(* CODESYS project xy_plotter.export

Project tree, tasks and I/O mapping:
  Device : CODESYS Control for Raspberry Pi 64 SL, CODESYS, order no. 2302000009, version 4.21.0.0
    application Application
      libraries: Standard, 3.5.22.0 (System); Net Base Services, * (CODESYS)
      task Main_OB1 (cyclic, interval t#4ms, priority 1) calls FB100_Logic_Call
      Drawing/
        global variables Drawing
      ESP Data/
        global variables RCV_ESP_Buffer
        global variables SND_ESP_Buffer
      HMI Data/
        global variables DB
      PLC data types/
        data type ESP_Cmd
        data type ESP_Coord
        data type ESP_Resp
        data type ESP_Zsw
        data type PLC_Contour
        data type PLC_Point
        data type TMR
        TCP/
          data type TCP_Con
          data type TCP_ESP_RCV
          data type TCP_ESP_SND
          data type TCP_Rcv
          data type TCP_Snd
      program FB100_Logic_Call [ST]
      function block FB200_TCP_ESP [ST]
      function block FB300_ESP_Cmd [ST]: AssignBit
      Symbols
    SoftMotion General Axis Pool
    GPIOs_A_B : GPIOs A/B, CODESYS, version 4.21.0.0
        unmapped channels: digital inputs (GPIO0..GPIO31), digital outputs (GPIO0..GPIO31)
    Onewire
    Camera device
      <Empty>
    SPI
    I²C
*)

// Device/Application/PLC data types/ESP_Cmd
TYPE ESP_Cmd :
	
STRUCT
    Stw         : UINT := 0;   // ESP32 control word
    PointFlags  : UINT := 0;   // Point command flags
    ContourNum  : UINT := 0;   // Contour number
    PointNum    : UINT := 0;   // Point number
    Speed       : UINT := 0;   // Movement speed
    Coord_X     : UINT := 0;   // Target X coordinate
    Coord_Y     : UINT := 0;   // Target Y coordinate
	
	ManMoveSpeed		: UINT := 0;	// Manual movement speed	
	
	TargetX         	: UINT := 0;   // Target X coordinate
	TargetY         	: UINT := 0;   // Target Y coordinate
	TargetMoveSpeed 	: UINT := 0;   // Target movement speed
		
END_STRUCT

END_TYPE

// Device/Application/PLC data types/ESP_Coord
TYPE ESP_Coord :
	
STRUCT
    X : REAL := 0.0;
    Y : REAL := 0.0;
END_STRUCT

END_TYPE

// Device/Application/PLC data types/ESP_Resp
TYPE ESP_Resp :

STRUCT
    ZSW_Byte1     : BYTE := 16#00;      // Status byte 1
    ZSW_Byte2     : BYTE := 16#00;      // Status byte 2
    NumExpected   : UINT := 0;          // Next expected point number
    LastContRcv   : UINT := 0;          // Last contour received
    LastContDone  : UINT := 0;          // Last contour completed
    CurrPoint     : UINT := 0;          // Current point number
    Coord_X       : UINT := 0;          // Current X coordinate
    Coord_Y       : UINT := 0;          // Current Y coordinate
    PointsInBuffer: UINT := 0;          // Number of points currently stored
    ErrorCode     : UINT := 0;          // ESP32 error code
	DrawingState  : USINT := 0;	    	// Running - 1, aborted - 2, finished - 3
END_STRUCT

END_TYPE

// Device/Application/PLC data types/ESP_Zsw
TYPE ESP_Zsw :
	
STRUCT
    RdyForRcvNewPnt 	: BOOL := FALSE;
    RdyForEn        	: BOOL := FALSE;
    Enabled         	: BOOL := FALSE;
    Off1            	: BOOL := FALSE;
    Off2            	: BOOL := FALSE;
    PenDn           	: BOOL := FALSE;
    RdyStartNewDrw  	: BOOL := FALSE;
    RdyContPrevDrw  	: BOOL := FALSE;
    DrwProccAct     	: BOOL := FALSE;
    SnsrHomeX       	: BOOL := FALSE;
    SnsrHomeY       	: BOOL := FALSE;
    SnsrLimitX      	: BOOL := FALSE;
    SnsrLimitY      	: BOOL := FALSE;
    MovingAuto      	: BOOL := FALSE;
    MovingHome      	: BOOL := FALSE;
    MovingManual    	: BOOL := FALSE;
END_STRUCT

END_TYPE

// Device/Application/PLC data types/PLC_Contour
TYPE PLC_Contour :

STRUCT
    RcvdByEsp    : BOOL := FALSE;   // Contour received by ESP32
    Done         : BOOL := FALSE;   // Contour drawing completed
    StartIndex   : UINT := 0;       // Start index of contour in point buffer
    PointCount   : UINT := 0;       // Number of points in contour
    CurrentPoint : UINT := 0;       // Current point number
END_STRUCT

END_TYPE

// Device/Application/PLC data types/PLC_Point
TYPE PLC_Point :
	
STRUCT
    CmdType : UINT := 0;     // Point command type
    Speed   : UINT := 0;     // Movement speed
    Coord_X : UINT := 0;     // Target X coordinate
    Coord_Y : UINT := 0;     // Target Y coordinate
END_STRUCT

END_TYPE

// Device/Application/PLC data types/TMR
TYPE TMR :

STRUCT
	IN : BOOL := FALSE;      // Timer enable input
    PT : TIME := T#0MS;      // Preset time
    Q  : BOOL := FALSE;      // Timer output
END_STRUCT

END_TYPE

// Device/Application/PLC data types/TCP/TCP_Con
TYPE TCP_Con :

STRUCT
    Req    		: BOOL;
    Done   		: BOOL;
    Busy   		: BOOL;
    Error  		: BOOL;
	ErrorID		: NBS.ERROR;
    Active		: BOOL;
	ConnBusy    : BOOL;
	ConnError   : BOOL;
	ConnErrorID : NBS.ERROR;
	Connected   : BOOL;
END_STRUCT

END_TYPE

// Device/Application/PLC data types/TCP/TCP_ESP_RCV
TYPE TCP_ESP_RCV :
	
STRUCT
	ResponseZswByte1       : BYTE;         		// ESP32 status word
	ResponseZswByte2       : BYTE;         		// ESP32 status word
    ResponseNumExpected    : UINT := 0;    		// Next expected point number
    ResponseLastContRcv    : UINT := 0;    		// Last contour received
    ResponseLastContDone   : UINT := 0;    		// Last contour completed
    ResponseCurrPoint      : UINT := 0;    		// Current point number
    ResponseCoord_X        : UINT := 0;   		// Current X coordinate
    ResponseCoord_Y        : UINT := 0;    		// Current Y coordinate
    ResponsePointsInBuffer : UINT := 0;    		// Number of points currently stored in buffer
    ResponseErrorCode      : UINT := 0;    		// ESP32 error code
	ResponseDrawingState   : USINT := 0;	    // Running - 1, aborted - 2, finished - 3
END_STRUCT

END_TYPE

// Device/Application/PLC data types/TCP/TCP_ESP_SND
TYPE TCP_ESP_SND :
	
STRUCT
	CommandStw        : UINT := 0;   			// ESP32 control word
    CommandPointFlags : UINT := 0;   			// Point command flags
    CommandContourNum : UINT := 0;   			// Contour number
    CommandPointNum   : UINT := 0;   			// Point number
    CommandSpeed      : UINT := 0;   			// Movement speed
    CommandCoord_X    : UINT := 0;   			// Target X coordinate
    CommandCoord_Y    : UINT := 0;   			// Target Y coordinate
	CommandManMoveSpeed		: UINT := 0;		// Manual movement speed	
	CommandTargetX         	: UINT := 0;   		// Target X coordinate
	CommandTargetY         	: UINT := 0;   		// Target Y coordinate
	CommandTargetMoveSpeed 	: UINT := 0;   		// Target movement speed
END_STRUCT

END_TYPE

// Device/Application/PLC data types/TCP/TCP_Rcv
TYPE TCP_Rcv :

STRUCT
    Req    		: BOOL;
	Ndr    		: BOOL;
    Done   		: BOOL;
    Busy   		: BOOL;
    Error  		: BOOL;
	ErrorID		: NBS.ERROR;
    Status		: WORD;
	Len			: UDINT;
END_STRUCT

END_TYPE

// Device/Application/PLC data types/TCP/TCP_Snd
TYPE TCP_Snd :

STRUCT
    Req    		: BOOL;
    Done   		: BOOL;
    Busy   		: BOOL;
    Error  		: BOOL;
	ErrorID		: NBS.ERROR;
    Status		: WORD;
	Len			: UDINT;
END_STRUCT

END_TYPE

// Device/Application/Drawing/Drawing
{attribute 'qualified_only'}
VAR_GLOBAL
	
	TotalNumbContours 	: UINT := 0;                    	// Total number of contours
    TotalNumbPoints   	: UINT := 0;                    	// Total number of points

    Contour 			: ARRAY[0..700] OF PLC_Contour;     // Contour data array
    Points  			: ARRAY[0..7000] OF PLC_Point;      // Point data array

END_VAR

// Device/Application/ESP Data/RCV_ESP_Buffer
{attribute 'qualified_only'}
VAR_GLOBAL
	
    TCP_ESP_RCV	: TCP_ESP_RCV;         		

END_VAR

// Device/Application/ESP Data/SND_ESP_Buffer
{attribute 'qualified_only'}
VAR_GLOBAL
	TCP_ESP_SND : TCP_ESP_SND;
	Default : TCP_ESP_SND;
END_VAR

// Device/Application/HMI Data/DB
{attribute 'qualified_only'}
VAR_GLOBAL
	
    RcvDataFromPC : BOOL := FALSE; 					// Receive new data from PC												
    AutoCmd : BOOL := FALSE;						// Start automatic operation
    MoveCmd : BOOL := TRUE;							// Enable move
    HomeCmd : BOOL := FALSE;						// Start homing sequence
	MoveToTargetCmd : BOOL := FALSE;				// Start moving to target (during manual mode)
    StopCmd : BOOL := TRUE;							// Stop current operation
    EstopCmd : BOOL := FALSE;						// Emergency stop command
    CleanCmd : BOOL := FALSE;						// Clear ESP32 point buffer
    
	ManualPenDn : BOOL := FALSE;					// Move pen to down position manually
    ManMoveNorth : BOOL := FALSE;					// Manual movement commands
    ManMoveNEast : BOOL := FALSE;
    ManMoveEast  : BOOL := FALSE;
    ManMoveSEast : BOOL := FALSE;
    ManMoveSouth : BOOL := FALSE;
    ManMoveSWest : BOOL := FALSE;
    ManMoveWest  : BOOL := FALSE;
    ManMoveNWest : BOOL := FALSE;
	ManMoveSpeed : INT := 1000;
	
	TargetX : INT := 0;								 // Move to point (during manual mode)
	TargetY : INT := 0;
	TargetMoveSpeed : INT := 1000;
	TargetPenDn : BOOL := FALSE;
	
END_VAR

// Device/Application/FB100_Logic_Call
PROGRAM FB100_Logic_Call

VAR
	TcpPcDone      : BOOL := FALSE;
    TcpPcDataSaved : BOOL := FALSE;	

    xDeleteDrwReq  : BOOL := FALSE;
    xDeleteDrwDone : BOOL := FALSE;
    xAckReq        : BOOL := FALSE;
    xAckReset      : BOOL := FALSE;

    xEspConnected  : BOOL := FALSE;
    xEspSendDone   : BOOL := FALSE;
    xEspReceiveNdr : BOOL := FALSE;
    xEspSendReq    : BOOL := FALSE;
    xEspReceiveReq : BOOL := FALSE;

    xEspHomeX      : BOOL := FALSE;
    xEspHomeY      : BOOL := FALSE;
	
	PlcHeartbeat   : UDINT := 0;
	
	TargetReached  : BOOL := FALSE;
	
	EspCommLostTimer 	: TON;
	EspCommLost 		: BOOL := FALSE;
	
	FB300_ESP_Cmd : FB300_ESP_Cmd;
	FB200_TCP_ESP : FB200_TCP_ESP;
END_VAR

VAR CONSTANT
    RcvPcBufferSize : INT := 500;
    DrwContourSize  : INT := 500;
    DrwPointSize    : INT := 7000;
END_VAR


// pc: 192.168.0.100
// plc: 192.168.0.254
// esp: 192.168.0.154

// Plc Heartbit for Ignition
PlcHeartbeat := PlcHeartbeat + 2;

// Reset the homing command when automatic mode is active or both axes have reached their home positions
IF DB.AutoCmd OR (xEspHomeX AND xEspHomeY) THEN
	DB.HomeCmd := FALSE;
END_IF;

IF RCV_ESP_Buffer.TCP_ESP_RCV.ResponseLastContDone >= Drawing.TotalNumbContours THEN
	DB.AutoCmd := FALSE;
END_IF

// Reset the target moving command when both axes have reached their positions
TargetReached := ABS(UINT_TO_INT(RCV_ESP_Buffer.TCP_ESP_RCV.ResponseCoord_X) - DB.TargetX * 100) <= 1 AND ABS(UINT_TO_INT(RCV_ESP_Buffer.TCP_ESP_RCV.ResponseCoord_Y) - DB.TargetY * 100) <= 1;

IF DB.MoveToTargetCmd AND TargetReached THEN
    DB.MoveToTargetCmd := FALSE;
END_IF;

// Cancel automatic movement and homing when a stop command is active
IF DB.StopCmd THEN
	DB.AutoCmd := FALSE;
	DB.HomeCmd := FALSE;
	DB.MoveToTargetCmd := FALSE;
END_IF;

// Prepare commands and exchange drawing data with the ESP
FB300_ESP_Cmd(Enable := NOT DB.RcvDataFromPC,
              ContourTotalNum := Drawing.TotalNumbContours,
              PointsTotalNum := Drawing.TotalNumbPoints,
              TCP_Conn_Estab := xEspConnected,
              TCP_Snd_Done := xEspSendDone,
              TCP_Rcv_Ndr := xEspReceiveNdr,
			  ConnLost := EspCommLost,
              TCP_Snd_Req => xEspSendReq,
              TCP_Rcv_Req => xEspReceiveReq,
			  SnsrHomeX => xEspHomeX,
              SnsrHomeY => xEspHomeY);
			  
// Manage the TCP connection and data exchange between the PLC and ESP
FB200_TCP_ESP(Enable := NOT DB.RcvDataFromPC,
			  SndRequest  := xEspSendReq,
    		  RcvRequest  := xEspReceiveReq,
    		  Connected   => xEspConnected,
     		  SndDone     => xEspSendDone,
    		  RcvNdr      => xEspReceiveNdr);	

EspCommLostTimer(IN := NOT xEspReceiveNdr, PT := T#3S);
EspCommLost := EspCommLostTimer.Q;

END_PROGRAM

// Device/Application/FB300_ESP_Cmd
FUNCTION_BLOCK FB300_ESP_Cmd

VAR_INPUT
    Enable           		: BOOL;
    ContourTotalNum  		: UINT;
    PointsTotalNum   		: UINT;
    TCP_Conn_Estab   		: BOOL;
    TCP_Snd_Done     		: BOOL;
    TCP_Rcv_Ndr      		: BOOL;
	ConnLost				: BOOL;
END_VAR

VAR_OUTPUT
    TCP_Snd_Req     		: BOOL;
    TCP_Rcv_Req      		: BOOL;
    SavedPointNum    		: UINT;
    SnsrHomeX   : BOOL;
    SnsrHomeY   : BOOL;
END_VAR

VAR_IN_OUT
END_VAR

VAR
    SSW                 	: INT := 0;
    ErrPointNum         	: INT := 0;
    NewContDone         	: INT := 0;
    NewContRcvd         	: INT := 0;
    PrevContDone        	: INT := 0;
    PrevContRcvd        	: INT := 0;
    CurrNumExpected     	: UINT := 0;
    PrevNumExpected     	: UINT := 0;
    CurrContForSend     	: UINT := 0;
    PrevContForSend     	: UINT := 0;
    IsFirstPointOfContour 	: BOOL := FALSE;
    IsLastPointOfContour  	: BOOL := FALSE;
    CurrCoordEsp        	: ESP_Coord;
    EspZsw             		: ESP_Zsw;
    SAVE_TIMER         		: TON;
	RETRY_TIME				: TON;
	TonRetryQ 				: BOOL;
    SAVE_T             		: TMR;
	RtrigConnLost			: R_TRIG;
	
	DebugPointNum : UINT;
	DebugFirstPoint : BOOL;
	DebugPointFlags : UINT;
END_VAR

VAR_TEMP
    i_cntr 					: INT;
    j_cntr 					: INT;
END_VAR

VAR CONSTANT
END_VAR


SAVE_TIMER(IN := SSW > 1, PT := T#5S, Q => SAVE_T.Q);
RETRY_TIME(IN := Enable AND SSW = 5, PT := T#200MS, Q  => TonRetryQ);

// Reset state machine when disabled
IF NOT Enable THEN
	SSW := 0;
	PrevNumExpected := 0;
END_IF;

RtrigConnLost(CLK := ConnLost);

IF RtrigConnLost.Q THEN
	SSW := 0;
END_IF;

CASE SSW OF
		
	0:  // Initial state
		RCV_ESP_Buffer.TCP_ESP_RCV.ResponseZswByte1 := 0;
		RCV_ESP_Buffer.TCP_ESP_RCV.ResponseZswByte2 := 0;
		EspZsw.RdyForRcvNewPnt := FALSE;
		SND_ESP_Buffer.TCP_ESP_SND := SND_ESP_Buffer.Default;
		
		IF Enable THEN
			CurrContForSend := 1;
			PrevNumExpected := 0;
			SSW := 3;
		END_IF;
		
	1:  // Check whether the ESP is ready to receive a new point
		IF EspZsw.RdyForRcvNewPnt THEN
			CurrNumExpected := RCV_ESP_Buffer.TCP_ESP_RCV.ResponseNumExpected;
			
			// Reset contour number when ESP requests the first point of a new drawing
			IF CurrNumExpected = 1 THEN
				CurrContForSend := 1;
			END_IF;
			
			// ESP requests the first point or the next sequential point
			IF (CurrNumExpected = 1 OR CurrNumExpected = PrevNumExpected + 1) AND CurrNumExpected <= PointsTotalNum THEN
				SSW := 2;
			
				// Switch to the next contour when the requested point is outside the current contour range
				WHILE CurrNumExpected > Drawing.Contour[CurrContForSend].StartIndex + Drawing.Contour[CurrContForSend].PointCount - 1 AND CurrContForSend < Drawing.TotalNumbContours DO
					CurrContForSend := CurrContForSend + 1; 
				END_WHILE;
				
			// ESP received the last point
			ELSIF CurrNumExpected - 1 = PointsTotalNum THEN
				SSW := 3;
			
			// ESP is still requesting the previously sent point
			ELSIF CurrNumExpected = PrevNumExpected THEN
				SSW := 3;
			END_IF;
		ELSE
			// Send dummy values while still updating the control word.
			SND_ESP_Buffer.TCP_ESP_SND.CommandPointNum := 9999;
			SND_ESP_Buffer.TCP_ESP_SND.CommandSpeed := 9999;
			SND_ESP_Buffer.TCP_ESP_SND.CommandCoord_X := 9999;
			SND_ESP_Buffer.TCP_ESP_SND.CommandCoord_Y := 9999;
			AssignBit(Value := SND_ESP_Buffer.TCP_ESP_SND.CommandPointFlags, BitNumber := 0, State := FALSE);    // Clear bit 0
			AssignBit(Value := SND_ESP_Buffer.TCP_ESP_SND.CommandPointFlags, BitNumber := 1, State := FALSE);    // Clear bit 1
			AssignBit(Value := SND_ESP_Buffer.TCP_ESP_SND.CommandPointFlags, BitNumber := 2, State := FALSE);    // Clear bit 2
			SSW := 3;
		END_IF;
		
	2:  // Prepare point data in the send buffer
		
		// Point data
		SND_ESP_Buffer.TCP_ESP_SND.CommandPointNum := CurrNumExpected;                                  
		SND_ESP_Buffer.TCP_ESP_SND.CommandSpeed := Drawing.Points[CurrNumExpected].Speed;           
		SND_ESP_Buffer.TCP_ESP_SND.CommandCoord_X := Drawing.Points[CurrNumExpected].Coord_X;        
		SND_ESP_Buffer.TCP_ESP_SND.CommandCoord_Y := Drawing.Points[CurrNumExpected].Coord_Y;         
		
		// Detect the first and last point of the current contour
		IsFirstPointOfContour :=
			CurrNumExpected = Drawing.Contour[CurrContForSend].StartIndex;
		
		IsLastPointOfContour :=
			CurrNumExpected =
			Drawing.Contour[CurrContForSend].StartIndex
			+ Drawing.Contour[CurrContForSend].PointCount - 1;
		
		SND_ESP_Buffer.TCP_ESP_SND.CommandContourNum := CurrContForSend;
		
		AssignBit(Value := SND_ESP_Buffer.TCP_ESP_SND.CommandPointFlags, BitNumber := 0, State := IsLastPointOfContour);
		AssignBit(Value := SND_ESP_Buffer.TCP_ESP_SND.CommandPointFlags, BitNumber := 1, State := Drawing.Points[CurrNumExpected].CmdType <> 2);
		
		// Check whether this is the final point of the entire drawing
		AssignBit(Value := SND_ESP_Buffer.TCP_ESP_SND.CommandPointFlags, BitNumber := 2, State := CurrNumExpected = PointsTotalNum);
		
		IF Drawing.Points[CurrNumExpected].CmdType = 2 THEN
			DebugPointNum := CurrNumExpected;
			DebugFirstPoint := IsFirstPointOfContour;
			DebugPointFlags := SND_ESP_Buffer.TCP_ESP_SND.CommandPointFlags;
		END_IF;
		
		IF DB.CleanCmd THEN
			SND_ESP_Buffer.TCP_ESP_SND := SND_ESP_Buffer.Default;
		END_IF;
		
		SSW := 3;
		
	3:  // Prepare the control word
		
		SND_ESP_Buffer.TCP_ESP_SND.CommandManMoveSpeed := INT_TO_UINT(DB.ManMoveSpeed);
		SND_ESP_Buffer.TCP_ESP_SND.CommandTargetMoveSpeed := INT_TO_UINT(DB.TargetMoveSpeed);
		SND_ESP_Buffer.TCP_ESP_SND.CommandTargetX := INT_TO_UINT(DB.TargetX * 100);
		SND_ESP_Buffer.TCP_ESP_SND.CommandTargetY := INT_TO_UINT(DB.TargetY * 100);
		
		AssignBit(Value := SND_ESP_Buffer.TCP_ESP_SND.CommandStw, BitNumber := 0,  State := NOT DB.StopCmd);                                              // stop off1
		AssignBit(Value := SND_ESP_Buffer.TCP_ESP_SND.CommandStw, BitNumber := 1,  State := NOT DB.EstopCmd);                                             // estop off2
		AssignBit(Value := SND_ESP_Buffer.TCP_ESP_SND.CommandStw, BitNumber := 2,  State := DB.AutoCmd);                                                  // auto or manual move by hmi
		AssignBit(Value := SND_ESP_Buffer.TCP_ESP_SND.CommandStw, BitNumber := 3,  State := DB.MoveCmd);                                                  // move enable
		AssignBit(Value := SND_ESP_Buffer.TCP_ESP_SND.CommandStw, BitNumber := 4,  State := DB.HomeCmd);                                                  // home
		AssignBit(Value := SND_ESP_Buffer.TCP_ESP_SND.CommandStw, BitNumber := 5,  State := DB.CleanCmd);                                                 // clean buffer
		AssignBit(Value := SND_ESP_Buffer.TCP_ESP_SND.CommandStw, BitNumber := 6,  State := DB.ManualPenDn);                                              // manual mode: pen down
		AssignBit(Value := SND_ESP_Buffer.TCP_ESP_SND.CommandStw, BitNumber := 7,  State := DB.ManMoveEast OR DB.ManMoveNEast OR DB.ManMoveSEast);       // manual mode: X positive
		AssignBit(Value := SND_ESP_Buffer.TCP_ESP_SND.CommandStw, BitNumber := 8,  State := DB.ManMoveWest OR DB.ManMoveNWest OR DB.ManMoveSWest);       // manual mode: X negative
		AssignBit(Value := SND_ESP_Buffer.TCP_ESP_SND.CommandStw, BitNumber := 9,  State := DB.ManMoveNorth OR DB.ManMoveNEast OR DB.ManMoveNWest);      // manual mode: Y positive
		AssignBit(Value := SND_ESP_Buffer.TCP_ESP_SND.CommandStw, BitNumber := 10, State := DB.ManMoveSouth OR DB.ManMoveSEast OR DB.ManMoveSWest);      // manual mode: Y negative
		AssignBit(Value := SND_ESP_Buffer.TCP_ESP_SND.CommandStw, BitNumber := 11, State := DB.MoveToTargetCmd);      									 // target mode: start
		AssignBit(Value := SND_ESP_Buffer.TCP_ESP_SND.CommandStw, BitNumber := 12, State := DB.TargetPenDn);      										 // target mode: pen down
		
		// Continue with transmission when the TCP connection is established
		IF TCP_Conn_Estab THEN
			SSW := 4;
		ELSE
			SSW := 1;
		END_IF;
		
	4:  // Send point and control data
		IF TCP_Snd_Done THEN
			SSW := 5;
			
			// Store the last successfully sent point number
			IF EspZsw.RdyForRcvNewPnt AND SND_ESP_Buffer.TCP_ESP_SND.CommandPointNum <> 9999 THEN
				PrevNumExpected := SND_ESP_Buffer.TCP_ESP_SND.CommandPointNum;
			END_IF;
		END_IF;
		
	5:  // Wait for ESP response containing the next expected point number
		IF TCP_Rcv_Ndr THEN
			
			// Detect an unexpected jump in the requested point number
			IF RCV_ESP_Buffer.TCP_ESP_RCV.ResponseNumExpected > CurrNumExpected + 1 THEN
				ErrPointNum := ErrPointNum + 1;
			END_IF;
			
			NewContDone := UINT_TO_INT(RCV_ESP_Buffer.TCP_ESP_RCV.ResponseLastContDone);
			NewContRcvd := UINT_TO_INT(RCV_ESP_Buffer.TCP_ESP_RCV.ResponseLastContRcv);
			SSW := 6;
		ELSIF TonRetryQ THEN
			SSW := 4;	
		END_IF;
		
	6:  // Update ESP status word
		EspZsw.RdyForRcvNewPnt := RCV_ESP_Buffer.TCP_ESP_RCV.ResponseZswByte1.%X0;         // ready for rcv new point
		EspZsw.RdyForEn := RCV_ESP_Buffer.TCP_ESP_RCV.ResponseZswByte1.%X1;                // ready for switching on
		EspZsw.Enabled := RCV_ESP_Buffer.TCP_ESP_RCV.ResponseZswByte1.%X2;                 // enabled
		EspZsw.Off1 := RCV_ESP_Buffer.TCP_ESP_RCV.ResponseZswByte1.%X3;                    // off1
		EspZsw.Off2 := RCV_ESP_Buffer.TCP_ESP_RCV.ResponseZswByte1.%X4;                    // off2
		EspZsw.PenDn := RCV_ESP_Buffer.TCP_ESP_RCV.ResponseZswByte1.%X5;                   // pen down
		EspZsw.RdyContPrevDrw := RCV_ESP_Buffer.TCP_ESP_RCV.ResponseZswByte1.%X6;          // ready to continue drw
		EspZsw.RdyStartNewDrw := RCV_ESP_Buffer.TCP_ESP_RCV.ResponseZswByte1.%X7;          // ready to start new drw
		EspZsw.DrwProccAct := RCV_ESP_Buffer.TCP_ESP_RCV.ResponseZswByte2.%X0;             // drw in process
		EspZsw.SnsrHomeX := RCV_ESP_Buffer.TCP_ESP_RCV.ResponseZswByte2.%X1;               // sensor home x
		EspZsw.SnsrHomeY := RCV_ESP_Buffer.TCP_ESP_RCV.ResponseZswByte2.%X2;               // sensor home y
		EspZsw.SnsrLimitX := RCV_ESP_Buffer.TCP_ESP_RCV.ResponseZswByte2.%X3;              // sensor limit x
		EspZsw.SnsrLimitY := RCV_ESP_Buffer.TCP_ESP_RCV.ResponseZswByte2.%X4;              // sensor limit y
		EspZsw.MovingAuto := RCV_ESP_Buffer.TCP_ESP_RCV.ResponseZswByte2.%X5;              // auto move
		EspZsw.MovingHome := RCV_ESP_Buffer.TCP_ESP_RCV.ResponseZswByte2.%X6;              // homing move
		EspZsw.MovingManual := RCV_ESP_Buffer.TCP_ESP_RCV.ResponseZswByte2.%X7;            // manual move
		SSW := 7;
		
	7:  // Update contour status flags
		IF NewContDone > PrevContDone THEN                                        // Mark newly completed contours as done
			FOR i_cntr := PrevContDone + 1 TO NewContDone DO
				Drawing.Contour[i_cntr].Done := TRUE;
				
				// Periodically save the last completed point number
				IF i_cntr = NewContDone AND SAVE_T.Q THEN
					SavedPointNum := Drawing.Contour[i_cntr].StartIndex + Drawing.Contour[i_cntr].PointCount;
				END_IF;
			END_FOR;
		END_IF;
		
		// Mark newly received contours as received by the ESP
		IF NewContRcvd > PrevContRcvd THEN                                
			FOR i_cntr := PrevContRcvd + 1 TO NewContRcvd DO
				Drawing.Contour[i_cntr].RcvdByEsp := TRUE;
			END_FOR;
		END_IF;
		
		// Convert the current ESP coordinates to engineering units
		CurrCoordEsp.X := UINT_TO_REAL(RCV_ESP_Buffer.TCP_ESP_RCV.ResponseCoord_X) / 100;
		CurrCoordEsp.Y := UINT_TO_REAL(RCV_ESP_Buffer.TCP_ESP_RCV.ResponseCoord_Y) / 100;
		
		// Store contour status for comparison during the next cycle
		PrevContDone := NewContDone;
		PrevContRcvd := NewContRcvd;
		
		SSW := 1;
		
END_CASE;

// Generate TCP send and receive requests
TCP_Snd_Req := SSW = 4;
TCP_Rcv_Req := SSW = 5;
SnsrHomeX := EspZsw.SnsrHomeX;
SnsrHomeY := EspZsw.SnsrHomeY;

METHOD AssignBit

VAR_INPUT
    BitNumber : USINT;
    State     : BOOL;
END_VAR

VAR_IN_OUT
    Value : WORD;
END_VAR

IF State THEN
    Value := Value OR SHL(WORD#1, BitNumber);
ELSE
    Value := Value AND NOT SHL(WORD#1, BitNumber);
END_IF;
END_METHOD

END_FUNCTION_BLOCK

// Device/Application/FB200_TCP_ESP
{attribute 'no_assign'}
FUNCTION_BLOCK FB200_TCP_ESP

VAR_INPUT
	Enable 				: BOOL;
	SndRequest  		: BOOL;
    RcvRequest  		: BOOL;
END_VAR

VAR_IN_OUT
END_VAR

VAR_OUTPUT
	Connected 			: BOOL;
    SndDone   			: BOOL;
    RcvNdr    			: BOOL;
END_VAR

VAR
	SSW       			: INT := 0;
    OLD_SSW   			: INT := 0;
    TCP_Con   			: TCP_Con;
    Err       			: INT := 0;
    STEP_TIME 			: TON;
    RETRY_TIME			: TON;
    TonStepQ  			: BOOL;
    TonRetryQ 			: BOOL;
	
    RtrigEnable     	: R_TRIG;
    FtrigEnable     	: F_TRIG;
    ComOk     			: BOOL := FALSE;
    SendCntr  			: UINT := 0;
	
	TCP_Rcv   			: TCP_Rcv;
    TCP_Snd   			: TCP_Snd;
	
	fbClient 			: NBS.TCP_Client;
    fbRead   			: NBS.TCP_Read;
    fbWrite  			: NBS.TCP_Write;
	Connection			: NBS.IConnection;
	ipESP				: NBS.IPv4Address := (ipAddress := '192.168.0.154');
	
	TEST : BOOL;
END_VAR


// State timers
STEP_TIME(IN := SSW = 3, PT := T#5000MS, Q  => TonStepQ);
RETRY_TIME(IN := NOT TCP_Rcv.Ndr AND SSW > 0 AND SSW < 3, PT := T#5100MS, Q  => TonRetryQ);

// Detect communication enable and disable edges //
RtrigEnable(CLK := Enable);
FtrigEnable(CLK := Enable);

// Disconnect on communication enable/disable event or retry timeout
IF RtrigEnable.Q OR FtrigEnable.Q OR TonRetryQ THEN
    SSW := 3;
END_IF;

// Default commands
TCP_Con.Req := FALSE;
TCP_Snd.Req := FALSE;
TCP_Rcv.Req := FALSE;

// State machine
CASE SSW OF

    0:  // Initial step
        IF Enable THEN
            SSW := 1;
        END_IF;

    1:  // Establish connection
        TCP_Con.Req := TRUE;

        IF TCP_Con.Active THEN
            SSW := 2;

        ELSIF TCP_Con.Error THEN
            Err := Err + 1;
			SSW := 3;
            // SSW := 4;
        END_IF;

	2:  // Connected

		TCP_Con.Req := TRUE;
		TCP_Snd.Req := SndRequest;
		TCP_Rcv.Req := RcvRequest;
	
		IF TCP_Con.Error OR TCP_Snd.Error OR TCP_Rcv.Error THEN
			Err := Err + 1;
			SSW := 3;
		END_IF;
		
    3:  // Close connection
        TCP_Con.Req := FALSE;
        TCP_Snd.Req := FALSE;
        TCP_Rcv.Req := FALSE;
		
		IF TonStepQ THEN
            SSW := 0;
        END_IF;

ELSE

	SSW := 3;

END_CASE;

// TCP client
fbClient(
    xEnable       := TCP_Con.Req,
    xDone         => TCP_Con.Done,
    xBusy         => TCP_Con.Busy,
    xError        => TCP_Con.Error,
    eErrorID      => TCP_Con.ErrorID,
    itfIPAddress  := ipESP,
    uiPort        := 2001,
    xActive       => TCP_Con.Active,
    itfConnection => Connection
);

// Receive data from ESP
fbRead(
    xEnable       := TCP_Rcv.Req,
    xBusy         => TCP_Rcv.Busy,
    xError        => TCP_Rcv.Error,
    eErrorID      => TCP_Rcv.ErrorID,
    itfConnection := Connection,
    pData         := ADR(RCV_ESP_Buffer.TCP_ESP_RCV),
    udiSize       := SIZEOF(RCV_ESP_Buffer.TCP_ESP_RCV),
    xReady        => TCP_Rcv.Ndr,
    udiCount      => TCP_Rcv.Len
);

// Send data to ESP
fbWrite(
    xExecute      := TCP_Snd.Req,
    xDone         => TCP_Snd.Done,
    xBusy         => TCP_Snd.Busy,
    xError        => TCP_Snd.Error,
    eErrorID      => TCP_Snd.ErrorID,
    itfConnection := Connection,
    pData         := ADR(SND_ESP_Buffer.TCP_ESP_SND),
    udiSize       := SIZEOF(SND_ESP_Buffer.TCP_ESP_SND),
    udiCount      => TCP_Snd.Len
);

// Outputs for FB302_ESP_Cmd
Connected := TCP_Con.Active;
SndDone   := TCP_Snd.Done;
RcvNdr    := TCP_Rcv.Ndr;

END_FUNCTION_BLOCK
